// TIA Portal project "HydroSim" (V15.1)

(* hardware
DEVICE "S7-1200 station_1"  S7-1200 Station
   slot 0: "Rack_0"  S7-1200 Rack  Rack  V1.0
   slot 1: "PLC_1"  CPU 1214C DC/DC/DC  6ES7 214-1AG31-0XB0  V3.0
DEVICE "HMI_1"  KTP600 Basic color PN
   slot 0: "HMI_1"  KTP600 Basic color PN  6AV6 647-0AD11-3AX0  12.0.0.0
   slot 1: "HMI_RT_1"  KTP600 Basic color PN  6AV6 647-0AD11-3AX0  12.0.0.0
   slot 5: "HMI_1.IE_CP_1"  PROFINET Interface  12.0.0.0
      slot 1: "PROFINET Interface_1"  PROFINET Interface
         slot 1: "Port_1"  Port
*)

// ===== PLC "PLC_1"  CPU 1214C DC/DC/DC =====

VAR_GLOBAL   // PLC tag table "Default tag table"
   "ReadPump" AT %M27.0 : Bool;
   "ReadValve" AT %M27.1 : Bool;
   "ReadJunction" AT %M27.2 : Bool;
   "ReadTank" AT %M27.3 : Bool;
   "ReadPipe" AT %M27.4 : Bool;
END_VAR

VAR_GLOBAL   // PLC tag table "Zone 0"
   "Pump 1" AT %M0.0 : Bool;
   "Pump 2" AT %M0.1 : Bool;
   "Pump 3" AT %M0.2 : Bool;
   "Pump 4" AT %M0.3 : Bool;
   "Valve 1 Pre" AT %M0.4 : Bool;
   "Valve 2 Pre" AT %M0.5 : Bool;
   "Valve 3 Pre" AT %M0.6 : Bool;
   "Valve 4 Pre" AT %M0.7 : Bool;
   "Valve 1 Post" AT %M5.0 : Bool;
   "Valve 2 Post" AT %M5.1 : Bool;
   "Valve 3 Post" AT %M5.2 : Bool;
   "Valve 4 Post" AT %M5.3 : Bool;
END_VAR

VAR_GLOBAL   // PLC tag table "Zone 1"
   "Pump 11" AT %M11.0 : Bool;
   "Valve 11 Pre" AT %M11.1 : Bool;
   "Valve 11 Post" AT %M11.2 : Bool;
END_VAR

VAR_GLOBAL   // PLC tag table "Zone 2"
   "Pump 21" AT %M21.0 : Bool;
   "Valve 21 Pre" AT %M21.1 : Bool;
   "Valve 21 Post" AT %I21.2 : Bool;
END_VAR

VAR_GLOBAL   // PLC tag table "Zone 3"
   "Pump 31" AT %M31.0 : Bool;
   "Valve 31 Pre" AT %M31.1 : Bool;
   "Valve 31 Post" AT %M31.2 : Bool;
END_VAR

VAR_GLOBAL   // PLC tag table "Zone 4"
   "Pump 41" AT %M41.0 : Bool;
   "Valve 41 Pre" AT %M41.1 : Bool;
   "Valve 41 Post" AT %M41.2 : Bool;
END_VAR

TYPE "Pump"
   STRUCT
      Zone : Int;
      ID : Int;
      Status : Int;
      Flow : Real;
      Speed : Real;
      Quality : Real;
   END_STRUCT;
END_TYPE

TYPE "Valve"
   STRUCT
      Zone : Int;
      ID : Int;
      Status : Int;
      Flow : Real;
      Quality : Real;
   END_STRUCT;
END_TYPE

TYPE "Junction"
   STRUCT
      Zone : Int;
      ID : Int;
      Demand : Real;
      Quality : Real;
      Pressure : Real;
   END_STRUCT;
END_TYPE

TYPE "Tank"
   STRUCT
      Zone : Int;
      ID : Int;
      Level : Real;
      Quality : Real;
      Pressure : Real;
   END_STRUCT;
END_TYPE

TYPE "Pipe"
   STRUCT
      Zone : Int;
      ID : Int;
      Flow : Real;
      Quality : Real;
   END_STRUCT;
END_TYPE

DATA_BLOCK "Modbus_parameters"   // DB2
{ S7_Optimized_Access := 'TRUE' }
VERSION : 0.1
   VAR
      NDR : Bool;
      DR : Bool;
      ERROR : Bool;
      STATUS : Word;
      CONNECT : TCON_IP_v4;
   END_VAR
BEGIN
   CONNECT.InterfaceId := 64;
   CONNECT.ID := 16#1;
   CONNECT.LocalPort := 502;
END_DATA_BLOCK

DATA_BLOCK "MODBUS DATA"   // DB3
{ S7_Optimized_Access := 'FALSE' }
VERSION : 0.1
   VAR
      DATA_1 : Array[0..99] of Int;
   END_VAR
BEGIN
   DATA_1[18] := 0;   // Ready to read pump flag
   DATA_1[38] := 0;   // Ready to read valve flag
   // DATA_1[0] : Pump zone
   // DATA_1[1] : Pump Index / ID
   // DATA_1[2] : Status
   // DATA_1[3] : Flow integer (*100)
   // DATA_1[20] : Valve zone
   // DATA_1[21] : Valve Index / ID
   // DATA_1[22] : Status
   // DATA_1[23] : Flow integer (*100)
   // DATA_1[24] : Quality integer (*100)
   // DATA_1[40] : Junction zone
   // DATA_1[41] : Junction Index / ID
   // DATA_1[42] : Demand integer (*100)
   // DATA_1[60] : Tank zone
   // DATA_1[61] : Tank Index / ID
   // DATA_1[62] : Fill level integer (*100)
   // DATA_1[43] : Quality integer (*100)
   // DATA_1[63] : Quality integer (*100)
   // DATA_1[80] : Pipe zone
   // DATA_1[81] : Pipe Index / ID
   // DATA_1[82] : Flow integer (*100)
   // DATA_1[83] : Quality integer (*100)
   // DATA_1[4] : Speed integer (*100)
   // DATA_1[5] : Quality integer (*100)
   // DATA_1[44] : Pressure integer (*100)
   // DATA_1[64] : Pressure integer (*100)
   // DATA_1[98] : Ready to read pipe flag
   // DATA_1[78] : Ready to read tank flag
   // DATA_1[58] : Ready to read junction flag
END_DATA_BLOCK

DATA_BLOCK "DataStruct"   // DB4
{ S7_Optimized_Access := 'TRUE' }
VERSION : 0.1
   VAR
      Pumps : Array[0..7] of "Pump";
      Valves : Array[0..16] of "Valve";
      Tanks : Array[0..3] of "Tank";
      Junctions : Array[0..1] of "Junction";
      Pipes : Array[0..1] of "Pipe";
   END_VAR
BEGIN
   Valves[9].ID := 2;
   Valves[9].Zone := 1;
   Valves[8].ID := 1;
   Valves[8].Zone := 1;
   Valves[7].ID := 8;
   Valves[6].ID := 7;
   Valves[5].ID := 6;
   Valves[4].ID := 5;
   Valves[3].ID := 4;
   Valves[2].ID := 3;
   Valves[1].ID := 2;
   Valves[0].ID := 1;
   Tanks[3].ID := 4;
   Tanks[2].ID := 3;
   Tanks[1].ID := 2;
   Tanks[0].ID := 1;
   Pumps[0].ID := 1;
   Pumps[1].ID := 2;
   Pumps[2].ID := 3;
   Pumps[3].ID := 4;
   Pumps[4].Zone := 1;
   Pumps[4].ID := 1;
   Pumps[5].Zone := 2;
   Pumps[5].ID := 1;
   Pumps[6].Zone := 3;
   Pumps[6].ID := 1;
   Pumps[7].Zone := 4;
   Pumps[7].ID := 1;
   Valves[10].Zone := 2;
   Valves[10].ID := 1;
   Valves[11].Zone := 2;
   Valves[11].ID := 2;
   Valves[12].Zone := 3;
   Valves[12].ID := 1;
   Valves[13].Zone := 3;
   Valves[13].ID := 2;
   Valves[14].Zone := 4;
   Valves[14].ID := 1;
   Valves[15].Zone := 4;
   Valves[15].ID := 2;
   // Pumps[0] : Pump 0.1
   // Pumps[1] : Pump 0.2
   // Pumps[2] : Pump 0.3
   // Pumps[3] : Pump 0.4
   // Pumps[4] : Pump 1.1
   // Pumps[5] : Pump 2.1
   // Pumps[6] : Pump 3.1
   // Pumps[7] : Pump 4.1
   // Valves[0] : Valve 0.1 (before Tank 0.1)
   // Valves[1] : Valve 0.2 (after Tank 0.1)
   // Valves[2] : Valve 0.3 (before Tank 0.2)
   // Valves[3] : Valve 0.4 (after Tank 0.2)
   // Valves[4] : Valve 0.5 (before Tank 0.3)
   // Valves[5] : Valve 0.6 (after Tank 0.3)
   // Valves[6] : Valve 0.7 (before Tank 0.4)
   // Valves[7] : Valve 0.8 (after Tank 0.4)
   // Valves[8] : Valve 1.1 (before Pump 1.1)
   // Valves[9] : Valve 1.2 (after Pump 1.1)
   // Valves[10] : Valve 2.1 (before Pump 2.1)
   // Valves[11] : Valve 2.2 (after Pump 2.1)
   // Valves[12] : Valve 3.1 (before Pump 3.1)
   // Valves[13] : Valve 3.2 (after Pump 3.1)
   // Valves[14] : Valve 4.1 (before Pump 4.1)
   // Valves[15] : Valve 4.2 (after Pump 4.1)
   // Tanks[0] : Tank 0.1
   // Tanks[1] : Tank 0.2
   // Tanks[2] : Tank 0.3
   // Tanks[3] : Tank 0.4
   // Valves[16] : Valve 0.0 (after reservoir)
END_DATA_BLOCK

FUNCTION "PumpFunction" : Void   // FC1, SCL
{ S7_Optimized_Access := 'TRUE' }
VERSION : 0.1
   VAR_INPUT
      Zone : Int;
      ID : Int;
      Status : Int;
      Flow : Int;
      Speed : Int;
      Quality : Int;
   END_VAR
   VAR_IN_OUT
      Pumps : Array[0..7] of "Pump";
      ReadFlag : Int;
   END_VAR
   VAR_TEMP
      i : UInt;   // Array index to select the pump to write to
   END_VAR
   // // Pumps[0] : Pump 0.1
   // // Pumps[1] : Pump 0.2
   // // Pumps[2] : Pump 0.3
   // // Pumps[3] : Pump 0.4
   // // Pumps[4] : Pump 1.1
   // // Pumps[5] : Pump 2.1
   // // Pumps[6] : Pump 3.1
   // // Pumps[7] : Pump 4.1
BEGIN
   IF #ReadFlag = 1 THEN
       CASE #Zone OF
           0:  // Statement zone 0
               CASE #ID OF
                   1:  // Statement Pump 0.1
                       #i := 0
                       ;
                   2:  // Statement Pump 0.2
                       #i := 1;
                       ;
                   3:  // Statement Pump 0.3
                       #i := 2;
                       ;
                   4:  // Statement Pump 0.4
                       #i := 3;
                       ;
                   ELSE
                       // ERROR
                       ;
               END_CASE;
               ;
           1:  // Statement zone 1
               CASE #ID OF
                   1:  // Statement Pump 1.1
                       #i := 4;
                       ;
                   ELSE
                       // ERROR
                       ;
               END_CASE;
               ;
           2:  // Statement zone 2
               CASE #ID OF
                   1:  // Statement Pump 2.1
                       #i := 5;
                       ;
                   ELSE
                       // ERROR
                       ;
               END_CASE;
               ;
           3:  // Statement zone 3
               CASE #ID OF
                   1:  // Statement Pump 3.1
                       #i := 6;
                       ;
                   ELSE
                       // ERROR
                       ;
               END_CASE;
               ;
           4:  // Statement zone 4
               CASE #ID OF
                   1:  // Statement Pump 4.1
                       #i := 7;
                       ;
                   ELSE
                       // ERROR
                       ;
               END_CASE;
               ;
           ELSE
               // ERROR
               ;
       END_CASE;
       #Pumps[#i].Status := #Status;
       #Pumps[#i].Flow := #Flow / 100.0;
       #Pumps[#i].Speed := #Speed / 100.0;
       #Pumps[#i].Quality := #Quality / 100.0;

       #ReadFlag := 0;
   END_IF;
END_FUNCTION

FUNCTION "ValveFunction" : Void   // FC2, SCL
{ S7_Optimized_Access := 'TRUE' }
VERSION : 0.1
   VAR_INPUT
      Zone : Int;
      ID : Int;
      Status : Int;
      Flow : Int;
      Quality : Int;
   END_VAR
   VAR_IN_OUT
      Valves : Array[0..16] of "Valve";
      ReadFlag : Int;
   END_VAR
   VAR_TEMP
      i : UInt;   // Array index to select the tank to write to
   END_VAR
   // // Valves[0] : Valve 0.1 (before Tank 0.1)
   // // Valves[1] : Valve 0.2 (after Tank 0.1)
   // // Valves[2] : Valve 0.3 (before Tank 0.2)
   // // Valves[3] : Valve 0.4 (after Tank 0.2)
   // // Valves[4] : Valve 0.5 (before Tank 0.3)
   // // Valves[5] : Valve 0.6 (after Tank 0.3)
   // // Valves[6] : Valve 0.7 (before Tank 0.4)
   // // Valves[7] : Valve 0.8 (after Tank 0.4)
   // // Valves[8] : Valve 1.1 (before Pump 1.1)
   // // Valves[9] : Valve 1.2 (after Pump 1.1)
   // // Valves[10] : Valve 2.1 (before Pump 2.1)
   // // Valves[11] : Valve 2.2 (after Pump 2.1)
   // // Valves[12] : Valve 3.1 (before Pump 3.1)
   // // Valves[13] : Valve 3.2 (after Pump 3.1)
   // // Valves[14] : Valve 4.1 (before Pump 4.1)
   // // Valves[15] : Valve 4.2 (after Pump 4.1)
   // // Valves[16] : Valve 0.0 (after reservoir)
BEGIN
   IF #ReadFlag = 1 THEN
       CASE #Zone OF
           0:  // Statement zone 0
               CASE #ID OF
                   0:  // Statement Valve 0.0
                       #i := 16;
                       ;
                   1:  // Statement Valve 0.1
                       #i := 0;
                       ;
                   2:  // Statement Valve 0.2
                       #i := 1;
                       ;
                   3:  // Statement Valve 0.3
                       #i := 2;
                       ;
                   4:  // Statement Valve 0.4
                       #i := 3;
                       ;
                   5:  // Statement Valve 0.5
                       #i := 4;
                       ;
                   6:  // Statement Valve 0.6
                       #i := 5;
                       ;
                   7:  // Statement Valve 0.7
                       #i := 6;
                       ;
                   8:  // Statement Valve 0.8
                       #i := 7;
                       ;
                   ELSE
                       // ERROR
                       ;
               END_CASE;
               ;
           1:  // Statement zone 1
               CASE #ID OF
                   1:  // Statement Valve 1.1
                       #i := 8;
                       ;
                   2:  // Statement Valve 1.2
                       #i := 9;
                       ;
                   ELSE
                       // ERROR
                       ;
               END_CASE;
               ;
           2:  // Statement zone 2
               CASE #ID OF
                   1:  // Statement Valve 2.1
                       #i := 10;
                       ;
                   2:  // Statement Valve 2.2
                       #i := 11;
                       ;
                   ELSE
                       // ERROR
                       ;
               END_CASE;
               ;
           3:  // Statement zone 3
               CASE #ID OF
                   1:  // Statement Valve 3.1
                       #i := 12;
                       ;
                   2:  // Statement Valve 3.2
                       #i := 13;
                       ;
                   ELSE
                       // ERROR
                       ;
               END_CASE;
               ;
           4:  // Statement zone 4
               CASE #ID OF
                   1:  // Statement Valve 4.1
                       #i := 14;
                       ;
                   2:  // Statement Valve 4.2
                       #i := 15;
                       ;
                   ELSE
                       // ERROR
                       ;
               END_CASE;
               ;
           ELSE
               // ERROR
               ;
       END_CASE;
       #Valves[#i].Status := #Status;
       #Valves[#i].Flow := #Flow / 100.0;
       #Valves[#i].Quality := #Quality / 100.0;

       #ReadFlag := 0;
   END_IF;
END_FUNCTION

FUNCTION "TankFunction" : Void   // FC3, SCL
{ S7_Optimized_Access := 'TRUE' }
VERSION : 0.1
   VAR_INPUT
      Zone : Int;
      ID : Int;
      Level : Int;
      Quality : Int;
      Pressure : Int;
   END_VAR
   VAR_IN_OUT
      Tanks : Array[0..3] of "Tank";
      ReadFlag : Int;
   END_VAR
   VAR_TEMP
      i : UInt;   // Array index to select the tank to write to
   END_VAR
BEGIN
   IF #ReadFlag = 1 THEN
       CASE #Zone OF
           0:  // Statement zone 0
               CASE #ID OF
                   1:  // Statement Tank 0.1
                       #i := 0;
                       ;
                   2:  // Statement Tank 0.2
                       #i := 1;
                       ;
                   3:  // Statement Tank 0.3
                       #i := 2;
                       ;
                   4:  // Statement Tank 0.4
                       #i := 3;
                       ;
                   ELSE
                       // ERROR
                       ;
               END_CASE;
               ;
           ELSE
               // ERROR
               ;
       END_CASE;
       #Tanks[#i].Level := #Level / 100.0;
       #Tanks[#i].Quality := #Quality / 100.0;
       #Tanks[#i].Pressure := #Pressure / 100.0;

       #ReadFlag := 0;
       ;
   END_IF;
END_FUNCTION

FUNCTION "JunctionFunction" : Void   // FC4, SCL
{ S7_Optimized_Access := 'TRUE' }
VERSION : 0.1
   VAR_INPUT
      Zone : Int;
      ID : Int;
      Demand : Int;
      Quality : Int;
      Pressure : Int;
   END_VAR
   VAR_IN_OUT
      Junctions : Array[0..1] of "Junction";
      ReadFlag : Int;
   END_VAR
   VAR_TEMP
      i : UInt;   // Array index to select the junction to write to
   END_VAR
BEGIN
   IF #ReadFlag = 1 THEN
       CASE #Zone OF
           0:  // Statement zone 0
               CASE #ID OF
                   1:  // Statement Junction 0.1
                       //#i := 0;
                       ;
                   ELSE
                       // ERROR
                       ;
               END_CASE;
               ;
           1:  // Statement zone 1
               CASE #ID OF
                   1:  // Statement Junction 1.1
                       //#i := 1;
                       ;
                   ELSE
                       // ERROR
                       ;
               END_CASE;
               ;
           2:  // Statement zone 2
               CASE #ID OF
                   1:  // Statement Junction 2.1
                       //#i := 2;
                       ;
                   ELSE
                       // ERROR
                       ;
               END_CASE;
               ;
           3:  // Statement zone 3
               CASE #ID OF
                   1:  // Statement Junction 3.1
                       //#i := 3;
                       ;
                   ELSE
                       // ERROR
                       ;
               END_CASE;
               ;
           4:  // Statement zone 4
               CASE #ID OF
                   1:  // Statement Junction 4.1
                       //#i := 4;
                       ;
                   ELSE
                       // ERROR
                       ;
               END_CASE;
               ;
           ELSE
               // ERROR
               ;
       END_CASE;
       //#Junctions[#i].Demand := #Demand;
       //#Junctions[#i].Quality := #Quality;
       //#Junctions[#i].Pressure := #Pressure;

       #ReadFlag := 0;
   END_IF;
END_FUNCTION

FUNCTION "PipeFunction" : Void   // FC5, SCL
{ S7_Optimized_Access := 'TRUE' }
VERSION : 0.1
   VAR_INPUT
      Zone : Int;
      ID : Int;
      Flow : Int;
      Quality : Int;
   END_VAR
   VAR_IN_OUT
      Pipes : Array[0..1] of "Pipe";
      ReadFlag : Int;
   END_VAR
   VAR_TEMP
      i : UInt;   // Array index to select the junction to write to
   END_VAR
BEGIN
   IF #ReadFlag = 1 THEN
       CASE #Zone OF
           0:  // Statement zone 0
               CASE #ID OF
                   1:  // Statement Pipe 0.1
                       //#i := 0;
                       ;
                   ELSE
                       // ERROR
                       ;
               END_CASE;
               ;
           1:  // Statement zone 1
               CASE #ID OF
                   1:  // Statement Pipe 1.1
                       //#i := 1;
                       ;
                   ELSE
                       // ERROR
                       ;
               END_CASE;
               ;
           2:  // Statement zone 2
               CASE #ID OF
                   1:  // Statement Pipe 2.1
                       //#i := 2;
                       ;
                   ELSE
                       // ERROR
                       ;
               END_CASE;
               ;
           3:  // Statement zone 3
               CASE #ID OF
                   1:  // Statement Pipe 3.1
                       //#i := 3;
                       ;
                   ELSE
                       // ERROR
                       ;
               END_CASE;
               ;
           4:  // Statement zone 4
               CASE #ID OF
                   1:  // Statement Pipe 4.1
                       //#i := 4;
                       ;
                   ELSE
                       // ERROR
                       ;
               END_CASE;
               ;
           ELSE
               // ERROR
               ;
       END_CASE;
       #Pipes[#i].Flow := #Flow;
       #Pipes[#i].Quality := #Quality;

       #ReadFlag := 0;
   END_IF;
END_FUNCTION

ORGANIZATION_BLOCK "Main"   // OB1, FBD, ProgramCycle
TITLE = "Main Program Sweep (Cycle)"
{ S7_Optimized_Access := 'TRUE' }
VERSION : 0.1
   VAR CONSTANT
      defaultgate : String;
   END_VAR
BEGIN

REGION Network 1: Modbus Connection
   // Modbus server block to communicate over Modbus with the Raspberry Pi.
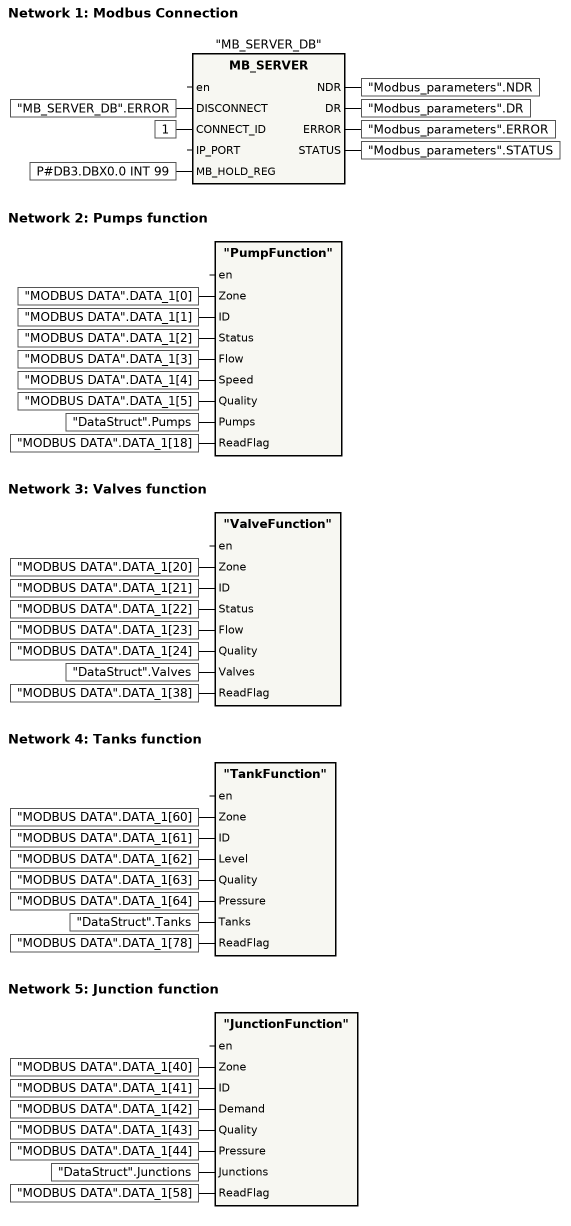
   "MB_SERVER_DB"(DISCONNECT := "MB_SERVER_DB".ERROR,   // MB_SERVER
                  CONNECT_ID := 1,
                  MB_HOLD_REG := P#DB3.DBX0.0 INT 99,
                  NDR => "Modbus_parameters".NDR,
                  DR => "Modbus_parameters".DR,
                  ERROR => "Modbus_parameters".ERROR,
                  STATUS => "Modbus_parameters".STATUS);
END_REGION

REGION Network 2: Pumps function
   // Function that reads the data from the Modbus server and copies the data to the right Pump UDT.
   "PumpFunction"(Zone := "MODBUS DATA".DATA_1[0],
                  ID := "MODBUS DATA".DATA_1[1],
                  Status := "MODBUS DATA".DATA_1[2],
                  Flow := "MODBUS DATA".DATA_1[3],
                  Speed := "MODBUS DATA".DATA_1[4],
                  Quality := "MODBUS DATA".DATA_1[5],
                  Pumps := "DataStruct".Pumps,
                  ReadFlag := "MODBUS DATA".DATA_1[18]);
END_REGION

REGION Network 3: Valves function
   // Function that reads the data from the Modbus server and copies the data to the right Valve UDT.
   "ValveFunction"(Zone := "MODBUS DATA".DATA_1[20],
                   ID := "MODBUS DATA".DATA_1[21],
                   Status := "MODBUS DATA".DATA_1[22],
                   Flow := "MODBUS DATA".DATA_1[23],
                   Quality := "MODBUS DATA".DATA_1[24],
                   Valves := "DataStruct".Valves,
                   ReadFlag := "MODBUS DATA".DATA_1[38]);
END_REGION

REGION Network 4: Tanks function
   // Function that reads the data from the Modbus server and copies the data to the right Tank UDT.
   "TankFunction"(Zone := "MODBUS DATA".DATA_1[60],
                  ID := "MODBUS DATA".DATA_1[61],
                  Level := "MODBUS DATA".DATA_1[62],
                  Quality := "MODBUS DATA".DATA_1[63],
                  Pressure := "MODBUS DATA".DATA_1[64],
                  Tanks := "DataStruct".Tanks,
                  ReadFlag := "MODBUS DATA".DATA_1[78]);
END_REGION

REGION Network 5: Junction function
   // Function that reads the data from the Modbus server and copies the data to the right Junction UDT.
   "JunctionFunction"(Zone := "MODBUS DATA".DATA_1[40],
                      ID := "MODBUS DATA".DATA_1[41],
                      Demand := "MODBUS DATA".DATA_1[42],
                      Quality := "MODBUS DATA".DATA_1[43],
                      Pressure := "MODBUS DATA".DATA_1[44],
                      Junctions := "DataStruct".Junctions,
                      ReadFlag := "MODBUS DATA".DATA_1[58]);
END_REGION

REGION Network 6: Pipe function
   // Function that reads the data from the Modbus server and copies the data to the right Pipe UDT.
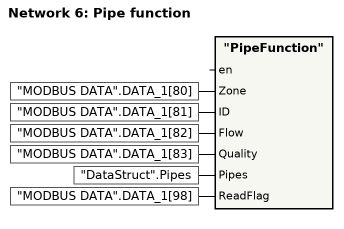
   "PipeFunction"(Zone := "MODBUS DATA".DATA_1[80],
                  ID := "MODBUS DATA".DATA_1[81],
                  Flow := "MODBUS DATA".DATA_1[82],
                  Quality := "MODBUS DATA".DATA_1[83],
                  Pipes := "DataStruct".Pipes,
                  ReadFlag := "MODBUS DATA".DATA_1[98]);
END_REGION
END_ORGANIZATION_BLOCK

(* ===== HMI "HMI_RT_1" =====
system functions are stored by id; their names below are inferred from use
connection "HMI_Connection_1": ETHERNET, SMART_S7_1200_OMS

HMI tags "Default tag table"
   "Tag_ScreenNumber" : UInt, internal
   "Pump 1" : Bool = PLC "Pump 1" AT %M0.0, 1 s
   "Pump 2" : Bool = PLC "Pump 2" AT %M0.1, 1 s
   "Pump 4" : Bool = PLC "Pump 4" AT %M0.3, 1 s
   "Pump 3" : Bool = PLC "Pump 3" AT %M0.2, 1 s
   "Valve 1 Post" : Bool = PLC "Valve 1 Post" AT %M5.0, 1 s
   "Valve 4 Post" : Bool = PLC "Valve 4 Post" AT %M5.3, 1 s
   "Valve 3 Post" : Bool = PLC "Valve 3 Post" AT %M5.2, 1 s
   "Valve 2 Post" : Bool = PLC "Valve 2 Post" AT %M5.1, 1 s
   "Valve 1 Pre" : Bool = PLC "Valve 1 Pre" AT %M0.4, 1 s
   "Valve 3 Pre" : Bool = PLC "Valve 3 Pre" AT %M0.6, 1 s
   "Valve 4 Pre" : Bool = PLC "Valve 4 Pre" AT %M0.7, 1 s
   "Valve 2 Pre" : Bool = PLC "Valve 2 Pre" AT %M0.5, 1 s
   "Pump 11" : Bool = PLC "Pump 11" AT %M11.0, 1 s
   "Valve 11 Pre" : Bool = PLC "Valve 11 Pre" AT %M11.1, 1 s
   "Valve 11 Post" : Bool = PLC "Valve 11 Post" AT %M11.2, 1 s
   "Valve 21 Pre" : Bool = PLC "Valve 21 Pre" AT %M21.1, 1 s
   "Pump 21" : Bool = PLC "Pump 21" AT %M21.0, 1 s
   "Valve 21 Post" : Bool = PLC "Valve 21 Post" AT %I21.2, 1 s
   "Valve 31 Pre" : Bool = PLC "Valve 31 Pre" AT %M31.1, 1 s
   "Pump 31" : Bool = PLC "Pump 31" AT %M31.0, 1 s
   "Valve 31 Post" : Bool = PLC "Valve 31 Post" AT %M31.2, 1 s
   "Valve 41 Pre" : Bool = PLC "Valve 41 Pre" AT %M41.1, 1 s
   "Pump 41" : Bool = PLC "Pump 41" AT %M41.0, 1 s
   "Valve 41 Post" : Bool = PLC "Valve 41 Post" AT %M41.2, 1 s
   "DataStruct_Pumps[0].Status" : Int = PLC DataStruct.Pumps[0].Status, 1 s
   "DataStruct_Pumps[1].Status" : Int = PLC DataStruct.Pumps[1].Status, 1 s
   "DataStruct_Pumps[3].Status" : Int = PLC DataStruct.Pumps[3].Status, 1 s
   "DataStruct_Pumps[2].Status" : Int = PLC DataStruct.Pumps[2].Status, 1 s
   "DataStruct_Valves[0].Status" : Int = PLC DataStruct.Valves[0].Status, 1 s
   "DataStruct_Valves[1].Status" : Int = PLC DataStruct.Valves[1].Status, 1 s
   "DataStruct_Valves[2].Status" : Int = PLC DataStruct.Valves[2].Status, 1 s
   "DataStruct_Valves[3].Status" : Int = PLC DataStruct.Valves[3].Status, 1 s
   "DataStruct_Valves[4].Status" : Int = PLC DataStruct.Valves[4].Status, 1 s
   "DataStruct_Valves[5].Status" : Int = PLC DataStruct.Valves[5].Status, 1 s
   "DataStruct_Valves[6].Status" : Int = PLC DataStruct.Valves[6].Status, 1 s
   "DataStruct_Valves[7].Status" : Int = PLC DataStruct.Valves[7].Status, 1 s
   "DataStruct_Pumps[4].Status" : Int = PLC DataStruct.Pumps[4].Status, 1 s
   "DataStruct_Valves[8].Status" : Int = PLC DataStruct.Valves[8].Status, 1 s
   "DataStruct_Valves[9].Status" : Int = PLC DataStruct.Valves[9].Status, 1 s
   "DataStruct_Pumps[5].Status" : Int = PLC DataStruct.Pumps[5].Status, 1 s
   "DataStruct_Valves[10].Status" : Int = PLC DataStruct.Valves[10].Status, 1 s
   "DataStruct_Valves[11].Status" : Int = PLC DataStruct.Valves[11].Status, 1 s
   "DataStruct_Pumps[6].Status" : Int = PLC DataStruct.Pumps[6].Status, 1 s
   "DataStruct_Valves[12].Status" : Int = PLC DataStruct.Valves[12].Status, 1 s
   "DataStruct_Valves[13].Status" : Int = PLC DataStruct.Valves[13].Status, 1 s
   "DataStruct_Pumps[7].Status" : Int = PLC DataStruct.Pumps[7].Status, 1 s
   "DataStruct_Valves[14].Status" : Int = PLC DataStruct.Valves[14].Status, 1 s
   "DataStruct_Valves[15].Status" : Int = PLC DataStruct.Valves[15].Status, 1 s
   "DataStruct_Tanks[0].Level" : Real = PLC DataStruct.Tanks[0].Level, 1 s
   "DataStruct_Tanks[2].Level" : Real = PLC DataStruct.Tanks[2].Level, 1 s
   "DataStruct_Valves[16].Status" : Int = PLC DataStruct.Valves[16].Status, 1 s

Template "Template_1" 320x240
   Button "Exit" at 266,202 size 52x37; TextOff 'Exit'; PictureOff "ExitRuntime_KTP600_Basic_color_PN"; PictureOn "ExitRuntime_KTP600_Basic_color_PN"
      on Release: StopRuntime(0)
   Button "Template_Button" at 213,202 size 52x37; TextOff 'Text'
   Button "Template_Button_1" at 160,202 size 52x37; TextOff 'Text'
   Button "Template_Button_2" at 107,202 size 52x37; TextOff 'Text'
   Button "Alarms" at 54,202 size 52x37; TextOff 'Alarms'; PictureOff "AlarmDisplay_KTP600_Basic_color_PN"; PictureOn "AlarmDisplay_KTP600_Basic_color_PN"
      on Release: function_ef3f5d25("Alarm window_Unacknowledged", -1)
   Button "Start screen" at 1,202 size 52x37; TextOff 'Start screen'; PictureOff "NavigateHome_KTP600_Basic_color_PN"; PictureOn "NavigateHome_KTP600_Basic_color_PN"
      on Release: ActivateScreen("HydroSim HMI", 0)
   SymbolicIOField "Symbolic_IO_Field_Screen" at 69,7 size 164x24; TextOff '0'; TextOn '1'; TextList "TextList_ScreenNames"
      ProcessValue <- "Tag_ScreenNumber"
      on Change: ActivateScreenByNumber("Tag_ScreenNumber", 0)
   DateTimeField "HmiScreenItemData" at 235,19 size 85x19
   DateTimeField "HmiScreenItemData_1" at 235,0 size 85x19
   GraphicView "Logo" at 0,0 size 67x38; Picture "Logo of HMI_1"

screen "HydroSim HMI" 320x240, template "Template_1"
   on GenerateScreen: SetTag("Tag_ScreenNumber", 1)
   TextField "HmiScreenItemData" at 32,109 size 256x17; Text 'Welcome to the HydroSim physical visualisation!'
   Button "Screen0" at 1,39 size 104x30; TextOff 'Zone 0'
      on Release: ActivateScreen("Zone 0", 0)
      on Click: ActivateScreen("Zone 0", 0)
   Button "Screen1" at 106,39 size 104x30; TextOff 'Zone 1'
      on Release: ActivateScreen("Zone 1", 0)
      on Click: ActivateScreen("Zone 1", 0)
   Button "Screen2" at 56,69 size 104x30; TextOff 'Zone 3'; TextOn 'Zone 2'
      on Release: ActivateScreen("Zone 3", 0)
      on Click: ActivateScreen("Zone 3", 0)
   Button "Screen3" at 160,69 size 104x30; TextOff 'Zone 4'; TextOn 'Zone 3'
      on Release: ActivateScreen("Zone 4", 0)
      on Click: ActivateScreen("Zone 4", 0)
   Button "Screen4" at 210,39 size 104x30; TextOff 'Zone 2'; TextOn 'Zone 4'
      on Release: ActivateScreen("Zone 2", 0)
      on Click: ActivateScreen("Zone 2", 0)

screen "Zone 0" 320x240, template "Template_1"
   on GenerateScreen: SetTag("Tag_ScreenNumber", 2)
   GraphicView "Graphic view_1" at 0,0 size 320x240; Picture "Zone0"
   Button "Back" at 0,210 size 104x30; TextOff 'Back'
      on Release: ActivateScreen("HydroSim HMI", 0)
   Circle "Circle_1" at 127,33 size 20x20
      Visibility <- "DataStruct_Pumps[0].Status"
   Rectangle "Rectangle_1" at 230,145 size 25x19
      Visibility <- "DataStruct_Valves[0].Status"
   Rectangle "Rectangle_2" at 204,145 size 25x19
      Visibility <- "DataStruct_Valves[2].Status"
   Rectangle "Rectangle_3" at 176,145 size 25x19
      Visibility <- "DataStruct_Valves[6].Status"
   Rectangle "Rectangle_4" at 148,145 size 25x19
      Visibility <- "DataStruct_Valves[4].Status"
   Rectangle "Rectangle_5" at 230,210 size 25x19
      Visibility <- "DataStruct_Valves[1].Status"
   Rectangle "Rectangle_6" at 204,210 size 25x19
      Visibility <- "DataStruct_Valves[3].Status"
   Rectangle "Rectangle_7" at 176,210 size 25x19
      Visibility <- "DataStruct_Valves[7].Status"
   Rectangle "Rectangle_8" at 148,210 size 25x19
      Visibility <- "DataStruct_Valves[5].Status"
   Circle "Circle_2" at 127,56 size 20x20
      Visibility <- "DataStruct_Pumps[1].Status"
   Circle "Circle_3" at 127,100 size 20x20
      Visibility <- "DataStruct_Pumps[3].Status"
   Circle "Circle_4" at 127,123 size 20x20
      Visibility <- "DataStruct_Pumps[2].Status"
   Bar "Bar_1" at 230,170 size 28x36; MinimumValue 0; MaximumValue 15
      ProcessValue <- "DataStruct_Tanks[0].Level"
   Bar "Bar_2" at 150,169 size 28x36; MinimumValue 0; MaximumValue 15
      ProcessValue <- "DataStruct_Tanks[2].Level"
   Rectangle "Rectangle_9" at 28,59 size 25x19
      Visibility <- "DataStruct_Valves[16].Status"

screen "Zone 1" 320x240, template "Template_1"
   on GenerateScreen: SetTag("Tag_ScreenNumber", 3)
   TextField "HmiScreenItemData" at 32,109 size 256x17; Text 'Screen1'
   GraphicView "Graphic view_1" at 0,0 size 320x240; Picture "Zone1"
   Button "Back" at 0,210 size 104x30; TextOff 'Back'
      on Release: ActivateScreen("HydroSim HMI", 0)
   Circle "Circle_1" at 84,168 size 20x20
      Visibility <- "DataStruct_Pumps[4].Status"
   Rectangle "Rectangle_8" at 114,174 size 25x19
      Visibility <- "DataStruct_Valves[9].Status"
   Rectangle "Rectangle_1" at 45,167 size 25x19
      Visibility <- "DataStruct_Valves[8].Status"

screen "Zone 2" 320x240, template "Template_1"
   on GenerateScreen: SetTag("Tag_ScreenNumber", 4)
   TextField "HmiScreenItemData" at 32,109 size 256x17; Text 'Screen2'
   GraphicView "Graphic view_1" at 0,0 size 320x240; Picture "Zone2"
   Button "Back" at 0,210 size 104x30; TextOff 'Back'
      on Release: ActivateScreen("HydroSim HMI", 0)
   Circle "Circle_1" at 84,168 size 20x20
      Visibility <- "DataStruct_Pumps[5].Status"
   Rectangle "Rectangle_8" at 114,174 size 25x19
      Visibility <- "DataStruct_Valves[11].Status"
   Rectangle "Rectangle_1" at 45,167 size 25x19
      Visibility <- "DataStruct_Valves[10].Status"

screen "Zone 3" 320x240, template "Template_1"
   on GenerateScreen: SetTag("Tag_ScreenNumber", 5)
   TextField "HmiScreenItemData" at 32,109 size 256x17; Text 'Screen3'
   GraphicView "Graphic view_1" at 0,0 size 320x239; Picture "Zone3"
   Button "Back" at 0,209 size 104x30; TextOff 'Back'
      on Release: ActivateScreen("HydroSim HMI", 0)
   Circle "Circle_1" at 82,67 size 20x20
      Visibility <- "DataStruct_Pumps[6].Status"
   Rectangle "Rectangle_8" at 113,75 size 25x19
      Visibility <- "DataStruct_Valves[13].Status"
   Rectangle "Rectangle_1" at 44,68 size 25x19
      Visibility <- "DataStruct_Valves[12].Status"

screen "Zone 4" 320x240, template "Template_1"
   on GenerateScreen: SetTag("Tag_ScreenNumber", 6)
   TextField "HmiScreenItemData" at 32,109 size 256x17; Text 'Screen4'
   GraphicView "Graphic view_1" at 0,0 size 320x240; Picture "Zone4"
   Button "Back" at 0,209 size 104x30; TextOff 'Back'
      on Release: ActivateScreen("HydroSim HMI", 0)
   Circle "Circle_1" at 68,55 size 20x20
      Visibility <- "DataStruct_Pumps[7].Status"
   Rectangle "Rectangle_8" at 96,61 size 25x19
      Visibility <- "DataStruct_Valves[15].Status"
   Rectangle "Rectangle_1" at 36,56 size 25x19
      Visibility <- "DataStruct_Valves[14].Status"
*)